(* IEC 61131-3 sources: llm-plc-st-eval/codesys/dobles/I6, 6 files *)

(* ---- 01_Correcta.st ---- *)
(* DOBLE DE PRUEBA I6/Correcta - NO ES CORPUS. Esperado: veredicto 1 *)
FUNCTION_BLOCK FB_Temperatura
VAR_INPUT
    rawTemp : INT;
END_VAR
VAR_OUTPUT
    tempC : REAL;
    enfriador : BOOL;
    almSensor : BOOL;
END_VAR
VAR
    almPrev : BOOL;
END_VAR
IF rawTemp < 0 OR rawTemp > 27648 THEN
    almSensor := TRUE;
    enfriador := FALSE;
ELSE
    almSensor := FALSE;
    tempC := INT_TO_REAL(rawTemp) / 27648.0 * 100.0;
    IF tempC >= 80.0 THEN
        enfriador := TRUE;
    ELSIF tempC <= 75.0 THEN
        enfriador := FALSE;
    END_IF
END_IF
END_FUNCTION_BLOCK

(* ---- 02_AlarmaNoApagaEnfriador.st ---- *)
(* DOBLE DE PRUEBA I6/AlarmaNoApagaEnfriador - NO ES CORPUS. Esperado: veredicto 2, falla en el paso 3 *)
FUNCTION_BLOCK FB_Temperatura
VAR_INPUT
    rawTemp : INT;
END_VAR
VAR_OUTPUT
    tempC : REAL;
    enfriador : BOOL;
    almSensor : BOOL;
END_VAR
VAR
    almPrev : BOOL;
END_VAR
IF rawTemp < 0 OR rawTemp > 27648 THEN
    almSensor := TRUE;
ELSE
    almSensor := FALSE;
    tempC := INT_TO_REAL(rawTemp) / 27648.0 * 100.0;
    IF tempC >= 80.0 THEN
        enfriador := TRUE;
    ELSIF tempC <= 75.0 THEN
        enfriador := FALSE;
    END_IF
END_IF
END_FUNCTION_BLOCK

(* ---- 03_SinHisteresis.st ---- *)
(* DOBLE DE PRUEBA I6/SinHisteresis - NO ES CORPUS. Esperado: veredicto 2, falla en el paso 2 *)
FUNCTION_BLOCK FB_Temperatura
VAR_INPUT
    rawTemp : INT;
END_VAR
VAR_OUTPUT
    tempC : REAL;
    enfriador : BOOL;
    almSensor : BOOL;
END_VAR
VAR
    almPrev : BOOL;
END_VAR
IF rawTemp < 0 OR rawTemp > 27648 THEN
    almSensor := TRUE;
    enfriador := FALSE;
ELSE
    almSensor := FALSE;
    tempC := INT_TO_REAL(rawTemp) / 27648.0 * 100.0;
    enfriador := tempC >= 80.0;
END_IF
END_FUNCTION_BLOCK

(* ---- 04_DivisionEntera.st ---- *)
(* DOBLE DE PRUEBA I6/DivisionEntera - NO ES CORPUS. Esperado: veredicto 2, falla en el paso 0 *)
FUNCTION_BLOCK FB_Temperatura
VAR_INPUT
    rawTemp : INT;
END_VAR
VAR_OUTPUT
    tempC : REAL;
    enfriador : BOOL;
    almSensor : BOOL;
END_VAR
VAR
    almPrev : BOOL;
END_VAR
IF rawTemp < 0 OR rawTemp > 27648 THEN
    almSensor := TRUE;
    enfriador := FALSE;
ELSE
    almSensor := FALSE;
    tempC := INT_TO_REAL(rawTemp / 27648 * 100);
    IF tempC >= 80.0 THEN
        enfriador := TRUE;
    ELSIF tempC <= 75.0 THEN
        enfriador := FALSE;
    END_IF
END_IF
END_FUNCTION_BLOCK

(* ---- 05_RangoSoloSuperior.st ---- *)
(* DOBLE DE PRUEBA I6/RangoSoloSuperior - NO ES CORPUS. Esperado: veredicto 2, falla en el paso 6 *)
FUNCTION_BLOCK FB_Temperatura
VAR_INPUT
    rawTemp : INT;
END_VAR
VAR_OUTPUT
    tempC : REAL;
    enfriador : BOOL;
    almSensor : BOOL;
END_VAR
VAR
    almPrev : BOOL;
END_VAR
IF rawTemp > 27648 THEN
    almSensor := TRUE;
    enfriador := FALSE;
ELSE
    almSensor := FALSE;
    tempC := INT_TO_REAL(rawTemp) / 27648.0 * 100.0;
    IF tempC >= 80.0 THEN
        enfriador := TRUE;
    ELSIF tempC <= 75.0 THEN
        enfriador := FALSE;
    END_IF
END_IF
END_FUNCTION_BLOCK

(* ---- 06_AlarmaEnclavada.st ---- *)
(* DOBLE DE PRUEBA I6/AlarmaEnclavada - NO ES CORPUS. Esperado: veredicto 2, falla en el paso 4 *)
FUNCTION_BLOCK FB_Temperatura
VAR_INPUT
    rawTemp : INT;
END_VAR
VAR_OUTPUT
    tempC : REAL;
    enfriador : BOOL;
    almSensor : BOOL;
END_VAR
VAR
    almPrev : BOOL;
END_VAR
almPrev := almSensor;
IF rawTemp < 0 OR rawTemp > 27648 THEN
    almSensor := TRUE;
    enfriador := FALSE;
ELSE
    almSensor := FALSE;
    tempC := INT_TO_REAL(rawTemp) / 27648.0 * 100.0;
    IF tempC >= 80.0 THEN
        enfriador := TRUE;
    ELSIF tempC <= 75.0 THEN
        enfriador := FALSE;
    END_IF
END_IF
almSensor := almSensor OR almPrev;
END_FUNCTION_BLOCK
